// TIA Portal V20 export
Screen "PN_DIAGNOSTIC_ALL"  1276x673
  ScreenItem "Line_Header_X0_Y64" at 0,64 size 1276x0  Type=HmiLine
  ScreenItem "Title_ScreenOverview_X390_Y2" at 390,2 size 500x30  Type=HmiTextBox
  ScreenItem "EA-Field_PN_IO_SYSTEM" at 725,35 size 60x25  Type=HmiIOField
  ScreenItem "PNIO-System" at 495,35 size 230x25  Type=HmiTextBox
  ScreenItem "PN-Diag_Reset" at 93,2 size 90x60  Type=HmiButton
  ScreenItem "PN-Diag_ReadNew" at 184,2 size 90x60  Type=HmiButton
  ScreenItem "Textfeld_1" at 292,8 size 95x22  Type=HmiTextBox
  ScreenItem "LED_1_Left_2" at 0,0 size 100x30  Type=HmiCircle
  ScreenItem "LED_1_Left_1" at 0,0 size 100x30  Type=HmiCircle
  ScreenItem "Textfeld_4" at 292,35 size 95x22  Type=HmiTextBox
  ScreenItem "permanentareaborderrectangle" at 0,0 size 0x0  Type=HmiRectangle
  ScreenItem "Button_Back" at 2,2 size 90x60  Type=HmiButton
  ScreenItem "PN-Diag_Counters" at 1093,2 size 90x60  Type=HmiButton
  ScreenItem "PN-Diag_LegendᆉY2" at 1184,2 size 90x60  Type=HmiButton
  ScreenItem "Rectangle_1" at 16,69 size 427x123  Type=HmiRectangle
  ScreenItem "LSicar_DeviceDiag_7" at 46,200 size 170x97  Type=HmiFaceplateContainer
  ScreenItem "LSicar_DeviceDiag_8" at 679,328 size 170x97  Type=HmiFaceplateContainer
  ScreenItem "LSicar_DeviceDiag_9" at 46,519 size 170x97  Type=HmiFaceplateContainer
  ScreenItem "LSicar_DeviceDiag_2" at 46,328 size 171x97  Type=HmiFaceplateContainer
  ScreenItem "LSicar_DeviceDiag_4" at 46,78 size 170x97  Type=HmiFaceplateContainer
  ScreenItem "LSicar_DeviceDiag_11" at 258,78 size 170x105  Type=HmiFaceplateContainer
  ScreenItem "LSicar_DeviceDiag_3" at 679,200 size 170x97  Type=HmiFaceplateContainer
  ScreenItem "LSicar_DeviceDiag_5" at 471,328 size 170x97  Type=HmiFaceplateContainer
  ScreenItem "LSicar_DeviceDiag_10" at 471,78 size 170x97  Type=HmiFaceplateContainer
  ScreenItem "LSicar_DeviceDiag_12" at 470,200 size 170x97  Type=HmiFaceplateContainer
  ScreenItem "LSicar_DeviceDiag_1" at 234,519 size 170x97  Type=HmiFaceplateContainer
  ScreenItem "LSicar_DeviceDiag_6" at 423,519 size 170x97  Type=HmiFaceplateContainer
  ScreenItem "LSicar_DeviceDiag_14" at 611,519 size 170x97  Type=HmiFaceplateContainer
  ScreenItem "LSicar_DeviceDiag_15" at 800,519 size 170x97  Type=HmiFaceplateContainer
  ScreenItem "LSicar_DeviceDiag_16" at 989,519 size 170x97  Type=HmiFaceplateContainer
  ScreenItem "Faceplate container_1" at 679,78 size 170x100  Type=HmiFaceplateContainer
  ScreenItem "LSicar_DeviceDiag_13" at 890,200 size 170x97  Type=HmiFaceplateContainer
  ScreenItem "线_18" at 410,638 size 120x0  Type=HmiLine
  ScreenItem "线_19" at 530,602 size 0x35  Type=HmiLine
  ScreenItem "线_43" at 410,153 size 0x485  Type=HmiLine
  ScreenItem "线_44" at 541,637 size 178x0  Type=HmiLine
  ScreenItem "线_45" at 540,601 size 0x35  Type=HmiLine
  ScreenItem "线_46" at 719,602 size 0x35  Type=HmiLine
  ScreenItem "线_47" at 730,637 size 178x0  Type=HmiLine
  ScreenItem "线_48" at 729,601 size 0x35  Type=HmiLine
  ScreenItem "线_49" at 908,602 size 0x35  Type=HmiLine
  ScreenItem "线_50" at 919,638 size 178x0  Type=HmiLine
  ScreenItem "线_51" at 918,602 size 0x35  Type=HmiLine
  ScreenItem "线_52" at 1097,603 size 0x35  Type=HmiLine
  ScreenItem "线_12" at 163,636 size 178x0  Type=HmiLine
  ScreenItem "线_13" at 162,601 size 0x35  Type=HmiLine
  ScreenItem "线_14" at 341,602 size 0x35  Type=HmiLine
  ScreenItem "线_7" at 245,152 size 0x332  Type=HmiLine
  ScreenItem "线_10" at 24,484 size 220x0  Type=HmiLine
  ScreenItem "线_11" at 246,153 size 101x0  Type=HmiLine
  ScreenItem "线_15" at 25,636 size 126x0  Type=HmiLine
  ScreenItem "线_16" at 153,601 size 0x35  Type=HmiLine
  ScreenItem "线_17" at 23,487 size 0x150  Type=HmiLine
  ScreenItem "线_8" at 234,139 size 0x306  Type=HmiLine
  ScreenItem "线_9" at 166,446 size 67x0  Type=HmiLine
  ScreenItem "线_25" at 165,411 size 0x34  Type=HmiLine
  ScreenItem "线_35" at 235,142 size 113x0  Type=HmiLine
  ScreenItem "线_5" at 144,283 size 0x27  Type=HmiLine
  ScreenItem "线_27" at 227,127 size 121x0  Type=HmiLine
  ScreenItem "线_28" at 225,128 size 0x183  Type=HmiLine
  ScreenItem "线_29" at 145,312 size 79x0  Type=HmiLine
  ScreenItem "线_4" at 155,139 size 60x0  Type=HmiLine
  ScreenItem "线_6" at 218,120 size 0x19  Type=HmiLine
  ScreenItem "线_26" at 219,119 size 129x0  Type=HmiLine
  ScreenItem "线_3" at 459,129 size 0x182  Type=HmiLine
  ScreenItem "线_20" at 412,129 size 45x0  Type=HmiLine
  ScreenItem "线_21" at 461,312 size 126x0  Type=HmiLine
  ScreenItem "线_22" at 589,279 size 0x33  Type=HmiLine
  ScreenItem "线_23" at 600,279 size 0x33  Type=HmiLine
  ScreenItem "线_30" at 601,312 size 197x0  Type=HmiLine
  ScreenItem "线_31" at 798,279 size 0x33  Type=HmiLine
  ScreenItem "线_32" at 809,279 size 0x32  Type=HmiLine
  ScreenItem "线_33" at 809,312 size 200x0  Type=HmiLine
  ScreenItem "线_34" at 1009,280 size 0x32  Type=HmiLine
  ScreenItem "线_40" at 601,442 size 197x0  Type=HmiLine
  ScreenItem "线_41" at 600,409 size 0x33  Type=HmiLine
  ScreenItem "线_42" at 798,408 size 0x33  Type=HmiLine
  ScreenItem "线_36" at 412,139 size 37x0  Type=HmiLine
  ScreenItem "线_37" at 450,140 size 0x300  Type=HmiLine
  ScreenItem "线_38" at 450,442 size 138x0  Type=HmiLine
  ScreenItem "线_39" at 589,409 size 0x33  Type=HmiLine
  ScreenItem "线_53" at 583,183 size 210x0  Type=HmiLine
  ScreenItem "线_54" at 582,152 size 0x30  Type=HmiLine
  ScreenItem "线_55" at 795,158 size 0x24  Type=HmiLine
  ScreenItem "线_24" at 411,117 size 55x1  Type=HmiLine
  ScreenItem "线_1" at 466,119 size 0x62  Type=HmiLine
  ScreenItem "线_2" at 466,182 size 101x0  Type=HmiLine
  ScreenItem "线_62" at 570,134 size 0x47  Type=HmiLine
  ScreenItem "线_63" at 570,135 size 5x0  Type=HmiLine
